Staubli VAL3: utAppearance.pjx

--- utAppearance.pjx ---
Parameters version=s8.8.3Cs9_BS1660 stackSize=5000 millimeterUnit=true
Program file=start.pgx
Program file=stop.pgx
Data file=utAppearance.dtx

--- utAppearance.dtx ---
public bool bVisibility

--- start.pgx ---
program start()
begin
end

--- stop.pgx ---
program stop()
begin
end
